TYPE ST_SoftKey :
STRUCT
	bIsPressed:	BOOL;
	eState:		E_ButtonState;
END_STRUCT
END_TYPE

(* stored: Version 1.1.0.1, ProductVersion 3.1.4024.9
   DUT ST_SoftKey: Id {1f340fa3-72e5-40ca-86ad-7830aeb40543} *)
